FUNCTION_BLOCK Prensa_Vibropac_HMI (* Service Interface Function Block Type *)
  (* Standard: 61499-2 *)
  (* Version 1.0, 19/10/2026, Hidryco, Hidryco, IHM do Prensa_Vibropac *)
  PACKAGE Hidryco.HidrycoLib;
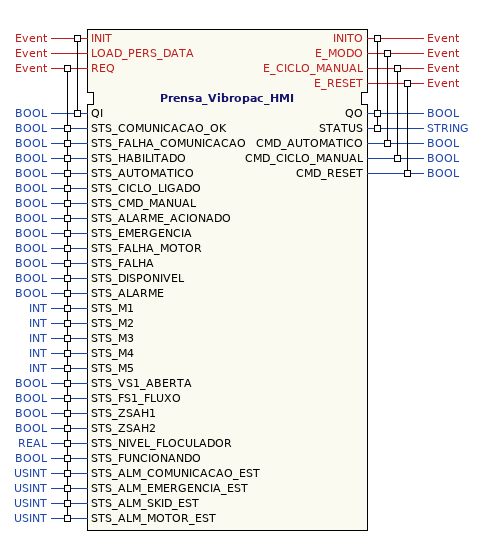
  EVENT_INPUT
    INIT WITH QI;
    LOAD_PERS_DATA; (* Reenvia os parametros persistentes *)
    REQ WITH STS_COMUNICACAO_OK, STS_FALHA_COMUNICACAO, STS_HABILITADO, STS_AUTOMATICO, STS_CICLO_LIGADO, STS_CMD_MANUAL, STS_ALARME_ACIONADO, STS_EMERGENCIA, STS_FALHA_MOTOR, STS_FALHA, STS_DISPONIVEL, STS_ALARME, STS_M1, STS_M2, STS_M3, STS_M4, STS_M5, STS_VS1_ABERTA, STS_FS1_FLUXO, STS_ZSAH1, STS_ZSAH2, STS_NIVEL_FLOCULADOR, STS_FUNCIONANDO, STS_ALM_COMUNICACAO_EST, STS_ALM_EMERGENCIA_EST, STS_ALM_SKID_EST, STS_ALM_MOTOR_EST; (* Atualizacao de status *)
  END_EVENT
  EVENT_OUTPUT
    INITO WITH QO, STATUS;
    E_MODO WITH CMD_AUTOMATICO;
    E_CICLO_MANUAL WITH CMD_CICLO_MANUAL;
    E_RESET WITH CMD_RESET;
  END_EVENT
  VAR_INPUT
    QI : BOOL;
    STS_COMUNICACAO_OK : BOOL; (* Comunicacao Modbus com o CLP do skid OK *)
    STS_FALHA_COMUNICACAO : BOOL; (* Falha de comunicacao com o CLP do skid *)
    STS_HABILITADO : BOOL; (* Instancia habilitada (FALSE = equipamento futuro) *)
    STS_AUTOMATICO : BOOL; (* Ciclo comandado pelo processo (automatico) *)
    STS_CICLO_LIGADO : BOOL; (* Comando de ciclo remoto ligado (4001 = 1) *)
    STS_CMD_MANUAL : BOOL; (* Comando manual de ciclo (modo manual) *)
    STS_ALARME_ACIONADO : BOOL; (* Alarme acionado no skid (4005) *)
    STS_EMERGENCIA : BOOL; (* Botao de emergencia do skid acionado (4006) *)
    STS_FALHA_MOTOR : BOOL; (* Algum motor do skid em falha *)
    STS_FALHA : BOOL; (* Skid em falha (alarme, emergencia ou motor) *)
    STS_DISPONIVEL : BOOL; (* Pode ser ligado pelo automatico agora *)
    STS_ALARME : BOOL; (* Algum alarme do skid *)
    STS_M1 : INT; (* Status M1 prensa (4007): 0 parado, 1 funcionando, 2 falha *)
    STS_M2 : INT; (* Status M2 motoredutor de limpeza (4008): 0 parado, 1 funcionando, 2 reverso, 3 falha *)
    STS_M3 : INT; (* Status M3 agitador do floculador (4009): 0 parado, 1 funcionando, 2 falha *)
    STS_M4 : INT; (* Status M4 bomba de agua (4010): 0 parado, 1 funcionando, 2 falha *)
    STS_M5 : INT; (* Status M5 compressor (4011): 0 parado, 1 funcionando, 2 falha *)
    STS_VS1_ABERTA : BOOL; (* Solenoide de limpeza VS1 aberta (4012) *)
    STS_FS1_FLUXO : BOOL; (* Chave de fluxo FS1 com fluxo (4013) *)
    STS_ZSAH1 : BOOL; (* Fim de curso frontal da limpeza atuado (4014) *)
    STS_ZSAH2 : BOOL; (* Fim de curso traseiro da limpeza atuado (4015) *)
    STS_NIVEL_FLOCULADOR : REAL; (* Nivel do tanque floculador LT1 (%) (4016, 0-1000) *)
    STS_FUNCIONANDO : BOOL; (* Prensa M1 funcionando *)
    STS_ALM_COMUNICACAO_EST : USINT; (* Estado do ALARM_BIT (0 normal, 1 ativo reconhecido, 2 ativo nao reconhecido, 3 saiu nao reconhecido, 4 ativo e saiu nao reconhecido) *)
    STS_ALM_EMERGENCIA_EST : USINT; (* Estado do ALARM_BIT (0 normal, 1 ativo reconhecido, 2 ativo nao reconhecido, 3 saiu nao reconhecido, 4 ativo e saiu nao reconhecido) *)
    STS_ALM_SKID_EST : USINT; (* Estado do ALARM_BIT (0 normal, 1 ativo reconhecido, 2 ativo nao reconhecido, 3 saiu nao reconhecido, 4 ativo e saiu nao reconhecido) *)
    STS_ALM_MOTOR_EST : USINT; (* Estado do ALARM_BIT (0 normal, 1 ativo reconhecido, 2 ativo nao reconhecido, 3 saiu nao reconhecido, 4 ativo e saiu nao reconhecido) *)
  END_VAR
  VAR_OUTPUT
    QO : BOOL; (* Event Output Qualifier *)
    STATUS : STRING; (* Service Status *)
    CMD_AUTOMATICO : BOOL; (* TRUE = automatico (ciclo pelo processo); persistente *)
    CMD_CICLO_MANUAL : BOOL; (* Manual: TRUE liga o ciclo remoto *)
    CMD_RESET : BOOL; (* Reset do skid (4002) e reconhecimento dos alarmes *)
  END_VAR
  SERVICE /
    SEQUENCE 
    END_SEQUENCE
  END_SERVICE
END_FUNCTION_BLOCK
